// TwinCAT 3 PLC project ExperimentSequencer
// ProgramVersion: 3.1.4026.22
// libraries:
//   Tc2_Standard, * (Beckhoff Automation GmbH)
//   Tc2_System, * (Beckhoff Automation GmbH)
// project tree:
//   DUTs/ E_SeqState.TcDUT
//   GVLs/ GVL_SEQ.TcGVL
//   POUs/ FB_ExperimentSequencerCore.TcPOU, PRG_ExperimentSequencer.TcPOU
//   / VirtualMotorTask.TcTTO
// (motion and I/O tree: see PLC project statemachinecontrol)
// real-time tasks:
//   TASK VirtualMotorTask: cycle T#125us, priority 1, ADS port 351
//   TASK StateTask: cycle T#10ms, priority 2, ADS port 355
// variable links:
//   ExperimentSequencer/ExperimentSequencer Instance <-> StateMachineControl/StateMachineControl Instance
//     VirtualMotorTask Inputs/GVL_SEQ.experimentActive <-> PlcTask Outputs/MAIN.experimentActiveOut
//     VirtualMotorTask Inputs/GVL_SEQ.resetReq <-> PlcTask Outputs/MAIN.resetOut
//     VirtualMotorTask Outputs/GVL_SEQ.playbackDone <-> PlcTask Inputs/MAIN.seqPlaybackDone
//   ExperimentSequencer/ExperimentSequencer Instance <-> ControllerCore/ControllerCore_Obj1 (Module1)
//     VirtualMotorTask Outputs/GVL_SEQ.ffValue <-> Inputs/ffValue
//     VirtualMotorTask Outputs/GVL_SEQ.refValue <-> Inputs/refValue
//   ExperimentSequencer/ExperimentSequencer Instance <-> DriverAdapter/DriverAdapter_Obj1 (Module1)
//     VirtualMotorTask Outputs/GVL_SEQ.distValue <-> Inputs/distValue
//     VirtualMotorTask Outputs/GVL_SEQ.playbackDone <-> Inputs/playbackDone
//   ExperimentSequencer/ExperimentSequencer Instance <-> ExperimentLogger/ExperimentLogger_Obj1 (Module1)
//     VirtualMotorTask Outputs/GVL_SEQ.distValue <-> Inputs/record/distValue
//     VirtualMotorTask Outputs/GVL_SEQ.ffValue <-> Inputs/record/ffValue
//     VirtualMotorTask Outputs/GVL_SEQ.playbackDone <-> Inputs/control/playbackDone
//     VirtualMotorTask Outputs/GVL_SEQ.refValue <-> Inputs/record/refValue

CONFIGURATION ExperimentSequencer
    RESOURCE PLC ON TwinCAT3
        TASK VirtualMotorTask(INTERVAL := T#125us, PRIORITY := 1);
        PROGRAM PRG_ExperimentSequencer WITH VirtualMotorTask : PRG_ExperimentSequencer;
    END_RESOURCE
END_CONFIGURATION

// ---- DUTs/E_SeqState.TcDUT
{attribute 'qualified_only'}
{attribute 'strict'}
TYPE E_SeqState :
(
    IDLE := 0,          (* Waiting. Outputs zeroed. *)
    PLAYING := 10,      (* Table playback active. *)
    COMPLETE := 20,     (* Playback complete, outputs held until rearm. *)
    FAULT := 90         (* Invalid input detected, reset edge required. *)
);
END_TYPE

// ---- GVLs/GVL_SEQ.TcGVL
{attribute 'qualified_only'}
VAR_GLOBAL CONSTANT
    N_REF_MAX : UDINT := 100000;
    N_FF_MAX : UDINT := 100000;
    N_DIST_MAX : UDINT := 100000;
END_VAR

VAR_GLOBAL
    {attribute 'linkalways'}
    refValue AT %Q* : LREAL := 0.0;

    {attribute 'linkalways'}
    ffValue AT %Q* : LREAL := 0.0;

    {attribute 'linkalways'}
    distValue AT %Q* : LREAL := 0.0;

    refTable : ARRAY[0..N_REF_MAX - 1] OF LREAL;
    ffTable : ARRAY[0..N_FF_MAX - 1] OF LREAL;
    distTable : ARRAY[0..N_DIST_MAX - 1] OF LREAL;
    tableLen : UDINT := 0;
    idx : UDINT := 0;
    repeatCount : UDINT := 1;
    trialIndex : UDINT := 0;

    {attribute 'linkalways'}
    resetReq AT %I* : BOOL := FALSE;

    {attribute 'linkalways'}
    experimentActive AT %I* : BOOL := FALSE;

    {attribute 'linkalways'}
    playbackDone AT %Q* : BOOL := FALSE;

    {attribute 'linkalways'}
    seqError AT %Q* : BOOL := FALSE;

    seqState : E_SeqState := E_SeqState.IDLE;
    tableLenClamped : UDINT := 0;
END_VAR

// ---- POUs/PRG_ExperimentSequencer.TcPOU
PROGRAM PRG_ExperimentSequencer
VAR
    tableIdxDint : DINT := 0;
    tableLenLocal : UDINT := 0;
    tableLenMaxLocal : UDINT := 0;
    refSample : LREAL := 0.0;
    ffSample : LREAL := 0.0;
    distSample : LREAL := 0.0;
    fbSequencerCore : FB_ExperimentSequencerCore;
END_VAR

tableLenMaxLocal := GVL_SEQ.N_REF_MAX;
IF GVL_SEQ.N_FF_MAX < tableLenMaxLocal THEN
    tableLenMaxLocal := GVL_SEQ.N_FF_MAX;
END_IF
IF GVL_SEQ.N_DIST_MAX < tableLenMaxLocal THEN
    tableLenMaxLocal := GVL_SEQ.N_DIST_MAX;
END_IF

tableLenLocal := GVL_SEQ.tableLen;
IF tableLenLocal > tableLenMaxLocal THEN
    tableLenLocal := tableLenMaxLocal;
END_IF
GVL_SEQ.tableLenClamped := tableLenLocal;

refSample := 0.0;
ffSample := 0.0;
distSample := 0.0;
IF fbSequencerCore.idx < tableLenLocal THEN
    tableIdxDint := UDINT_TO_DINT(fbSequencerCore.idx);
    refSample := GVL_SEQ.refTable[tableIdxDint];
    ffSample := GVL_SEQ.ffTable[tableIdxDint];
    distSample := GVL_SEQ.distTable[tableIdxDint];
END_IF

fbSequencerCore(
    resetRequest := GVL_SEQ.resetReq,
    experimentActive := GVL_SEQ.experimentActive,
    tableLen := tableLenLocal,
    repeatCount := GVL_SEQ.repeatCount,
    refSample := refSample,
    ffSample := ffSample,
    distSample := distSample
);

GVL_SEQ.refValue := fbSequencerCore.refValue;
GVL_SEQ.ffValue := fbSequencerCore.ffValue;
GVL_SEQ.distValue := fbSequencerCore.distValue;
GVL_SEQ.playbackDone := fbSequencerCore.playbackDone;
GVL_SEQ.seqError := fbSequencerCore.seqError;
GVL_SEQ.seqState := fbSequencerCore.seqState;
GVL_SEQ.idx := fbSequencerCore.idx;
GVL_SEQ.trialIndex := fbSequencerCore.trialIndex;

END_PROGRAM

// ---- POUs/FB_ExperimentSequencerCore.TcPOU
FUNCTION_BLOCK FB_ExperimentSequencerCore
VAR_INPUT
    resetRequest : BOOL;
    experimentActive : BOOL;
    tableLen : UDINT;
    repeatCount : UDINT;
    refSample : LREAL;
    ffSample : LREAL;
    distSample : LREAL;
END_VAR
VAR_OUTPUT
    refValue : LREAL := 0.0;
    ffValue : LREAL := 0.0;
    distValue : LREAL := 0.0;
    playbackDone : BOOL := FALSE;
    seqError : BOOL := FALSE;
    seqState : E_SeqState := E_SeqState.IDLE;
    idx : UDINT := 0;
    trialIndex : UDINT := 0;
END_VAR
VAR
    experimentActivePrev : BOOL := FALSE;
    resetRequestPrev : BOOL := FALSE;
    resetEdge : BOOL := FALSE;
    startEdge : BOOL := FALSE;
    zeroOutputsThisScan : BOOL := FALSE;
    resetProgressThisScan : BOOL := FALSE;
END_VAR

zeroOutputsThisScan := FALSE;
resetProgressThisScan := FALSE;
resetEdge := resetRequest AND NOT resetRequestPrev;
startEdge := experimentActive AND NOT experimentActivePrev;

IF resetEdge THEN
    resetProgressThisScan := TRUE;
    zeroOutputsThisScan := TRUE;
    seqState := E_SeqState.IDLE;

ELSE
    CASE seqState OF
        E_SeqState.IDLE:
            zeroOutputsThisScan := TRUE;

            IF startEdge THEN
                IF (tableLen = 0) OR (repeatCount = 0) THEN
                    seqState := E_SeqState.FAULT;
                ELSE
                    resetProgressThisScan := TRUE;
                    seqState := E_SeqState.PLAYING;
                END_IF
            END_IF

        E_SeqState.PLAYING:
            IF NOT experimentActive THEN
                resetProgressThisScan := TRUE;
                zeroOutputsThisScan := TRUE;
                seqState := E_SeqState.IDLE;
            ELSIF idx < tableLen THEN
                refValue := refSample;
                ffValue := ffSample;
                distValue := distSample;
                idx := idx + 1;

                IF idx >= tableLen THEN
                    IF trialIndex >= (repeatCount - 1) THEN
                        playbackDone := TRUE;
                        seqState := E_SeqState.COMPLETE;
                    ELSE
                        idx := 0;
                        trialIndex := trialIndex + 1;
                    END_IF
                END_IF
            END_IF

        E_SeqState.COMPLETE:
            IF NOT experimentActive THEN
                resetProgressThisScan := TRUE;
                zeroOutputsThisScan := TRUE;
                seqState := E_SeqState.IDLE;
            END_IF

        E_SeqState.FAULT:
            resetProgressThisScan := TRUE;
            zeroOutputsThisScan := TRUE;
    END_CASE
END_IF

IF resetProgressThisScan THEN
    idx := 0;
    trialIndex := 0;
END_IF
IF zeroOutputsThisScan THEN
    refValue := 0.0;
    ffValue := 0.0;
    distValue := 0.0;
    playbackDone := FALSE;
END_IF

seqError := (seqState = E_SeqState.FAULT);
experimentActivePrev := experimentActive;
resetRequestPrev := resetRequest;

END_FUNCTION_BLOCK
